// TIA Portal V20 export
TYPE "AXIS_FESTO_SIN_POS_TEL_111"
   STRUCT
      AXIS_TEL_111 : Struct
         SENDING : Struct
            MODE_POS : Int;   // JOG = 7 REALATIVE = 2 ABSOLUTNĚ = 1 HOMING = 4 / JOG = 7 RELATIVE = 2 ABSOLUTE = 1 HOMING = 4
            ENABLE_AXIS : Bool;   // ENABLE
            CANCEL_TRAVERSING : Bool;
            INTERMEDIATE_STOP : Bool;
            POSITIVE : Bool;
            NEGATIVE : Bool;
            JOG_1 : Bool;
            JOG_2 : Bool;
            FLI_REF : Bool;
            ACK_ERROR : Bool;
            EXECUTE_MODE : Bool;
            POSITION : DInt;
            VELOCITY : DInt;
            OVER_V : Int;
            OVER_ACC : Int;
            OVER_DEC : Int;
         END_STRUCT;
         READ : Struct
            AXIS_ENABLED : Bool;
            AXIS_POS_OK : Bool;
            AXIS_SP_FIXED : Bool;
            AXIS_REF : Bool;
            AXIS_WARN : Bool;
            AXIS_ERROR : Bool;
            LOCKOUT : Bool;
            ACT_VELOCITY : DInt;
            ACT_POSITION : DInt;
            ACT_MODE : Int;
            EPOS_ZSW_1 : Word;
            EPOS_ZSW_2 : Word;
            ACT_WARN : Word;
            ACT_FAULT : Word;
            ERROR : Bool;
            STATUS : Word;
            DIAGLD : Word;
         END_STRUCT;
      END_STRUCT;
   END_STRUCT;
END_TYPE
